// ── 10. Home ─────────────────────────────────────────────────────────────────
// Two-step home: MC_Direct sets the actual position, but does NOT raise the axis
// calibrated/Homed flag. MC_ForceCalibration then sets that flag (no motion, no
// position change). _homeCmd stays TRUE across both steps so all "home active"
// gates (jog/move blocking, fault) remain valid for the whole sequence.
IF NOT _homeCmd THEN
    _homeStep := 0;                     // sequence aborted elsewhere (stop/reset) → reset step
END_IF

// Step 1: set position
_mcHome(
    Axis       := Axis,
    Execute    := _homeCmd AND (_homeStep = 1),
    Position   := _homePosition,
    HomingMode := MC_Direct
);
IF _mcHome.Done AND (_homeStep = 1) THEN
    _homeStep          := 2;            // position set → now flag the axis as calibrated
    _dbgHomeDirectDone := TRUE;         // latch (diagnostic)
    // Retain the teach (section 10b) as an offset from the RAW encoder position, so it can be
    // re-applied after the NC restarts. Raw = the position before MC_Direct minus whatever offset
    // the running NC already applied.
    IF _retainHome THEN
        _homeOffset      := _homePosition - (_homeActAtStart - _ncOffsetApplied);
        _ncOffsetApplied := _homeOffset;
        _homeTaughtPos   := _homePosition;
        _homeTaught      := TRUE;
    END_IF
END_IF
IF _mcHome.Error THEN
    _homeCmd  := FALSE;
    _homeStep := 0;
    _lastMcErrorId := _mcHome.ErrorID;
    setFault(TRUE, CONCAT('Home error: ', UDINT_TO_STRING(_mcHome.ErrorID)));
END_IF
IF _homeStep > _dbgHomeMaxStep THEN _dbgHomeMaxStep := _homeStep; END_IF

// Step 2: set calibrated/Homed flag
_mcForceCal(
    Axis       := Axis,
    Execute    := _homeCmd AND (_homeStep = 2),
    HomingMode := MC_ForceCalibration
);
IF _mcForceCal.Done THEN
    _homeCmd        := FALSE;
    _homeStep       := 0;
    _dbgHomeCalDone := TRUE;            // latch (diagnostic)
END_IF
IF _mcForceCal.Error THEN
    _homeCmd         := FALSE;
    _homeStep        := 0;
    _dbgHomeCalError := TRUE;           // latch (diagnostic)
    _dbgHomeCalErrID := _mcForceCal.ErrorID;
    _lastMcErrorId := _mcForceCal.ErrorID;
    setFault(TRUE, CONCAT('Home cal error: ', UDINT_TO_STRING(_mcForceCal.ErrorID)));
END_IF

// ── 10b. Retained home ────────────────────────────────────────────────────────
// A taught home is kept (VAR PERSISTENT _homeTaught/_homeOffset) until the next teach — through
// PLC/NC restarts, activations and power cycles. MC_Direct only shifts the position inside the
// RUNNING NC, so after an NC restart (every activation) the axis reports the raw absolute-encoder
// position and is not homed. Once per PLC start, after the axis IO has been valid for 1 s (never
// act on a 0 read before EtherCAT is up), check the NC:
//   - not homed → the NC restarted and dropped the offset: MC_SetPosition(raw + offset), then
//                 MC_ForceCalibration. No motion and no enable needed.
//   - homed     → only the PLC restarted; the running NC still carries the offset: do nothing.
// Requires an ABSOLUTE encoder (cfgRetainHome := FALSE on an incremental one) and an NC encoder
// config that does not set the calibration flag by itself at startup.
_homeRestoreDelay(
    IN := _retainHome AND NOT _homeRestoreChecked
          AND NOT Axis.NcToPlc.StateDWord.30      // IoDataInvalid (StateDWord is a plain DWORD in Tc2_MC2)
          AND NOT Axis.NcToPlc.StateDWord.28      // DriveDeviceError
          AND NOT Axis.Status.Error,
    PT := T#1S
);
IF _homeRestoreDelay.Q THEN
    _homeRestoreChecked := TRUE;
    IF Axis.Status.Homed THEN
        _ncOffsetApplied := SEL(_homeTaught, 0.0, _homeOffset);
    ELSIF _homeTaught AND NOT _homeCmd AND NOT _externalControl THEN
        _ncOffsetApplied   := 0.0;
        _homeRestoreTarget := Axis.NcToPlc.ActPos + _homeOffset;
        _homeRestoreStep   := 1;
    END_IF
END_IF

_mcRestorePos(
    Axis     := Axis,
    Execute  := (_homeRestoreStep = 1),
    Position := _homeRestoreTarget,
    Mode     := FALSE                   // absolute
);
IF _mcRestorePos.Done AND (_homeRestoreStep = 1) THEN
    _ncOffsetApplied := _homeOffset;
    _homeRestoreStep := 2;
END_IF
IF _mcRestorePos.Error THEN
    _homeRestoreStep := 0;
    _lastMcErrorId := _mcRestorePos.ErrorID;
    setFault(TRUE, CONCAT('Home restore error: ', UDINT_TO_STRING(_mcRestorePos.ErrorID)));
END_IF

_mcRestoreCal(
    Axis       := Axis,
    Execute    := (_homeRestoreStep = 2),
    HomingMode := MC_ForceCalibration
);
IF _mcRestoreCal.Done THEN
    _homeRestoreStep := 0;
END_IF
IF _mcRestoreCal.Error THEN
    _homeRestoreStep := 0;
    _lastMcErrorId := _mcRestoreCal.ErrorID;
    setFault(TRUE, CONCAT('Home restore cal error: ', UDINT_TO_STRING(_mcRestoreCal.ErrorID)));
END_IF

// ── 11. Move execution state machine ──────────────────────────────────────────
// _moveExecState: 0=idle, 1=one-scan-abort (all Execute FALSE), 2=executing
// While yielded to an external coordinator (e.g. fb_CamCoupler), keep the state machine idle
// so every move block is driven Execute:=FALSE and never fights the external coupling.
IF _externalControl THEN
    _moveExecState := 0;
END_IF
// Arm new move request (set by cmdStart)
IF _startMoveReq AND NOT _stopCmd AND NOT _externalControl THEN
    _startMoveReq     := FALSE;
    _currentMoveIndex := _pendingIndex;
    _activeMoveMode   := _pendingMode;
    stsMoveDone       := FALSE;
    _haltCmd          := FALSE;
    _jogPositive      := FALSE;
    _jogNegative      := FALSE;
    IF _moveExecState = 2 THEN
        _moveExecState := 1; // one clear scan before rising edge on new block
    ELSE
        _moveExecState := 2;
    END_IF
END_IF

CASE _moveExecState OF

    0, 1: // Idle or abort-scan: drive all move blocks with Execute FALSE
        _mcMoveAbs(Axis := Axis, Execute := FALSE, Position := 0.0,     Velocity := 1.0, Acceleration := 1.0, Deceleration := 1.0, Jerk := 0.0);
        _mcMoveRel(Axis := Axis, Execute := FALSE, Distance := 0.0,     Velocity := 1.0, Acceleration := 1.0, Deceleration := 1.0, Jerk := 0.0);
        _mcMoveVel(Axis := Axis, Execute := FALSE);
        _mcTorque( Axis := Axis, Execute := FALSE);
        _mcMoveMod(Axis := Axis, Execute := FALSE);
        IF _moveExecState = 1 THEN
            _moveExecState := 2; // transition to executing next scan
        END_IF

    2: // Executing - drive only the active mode block; others get Execute FALSE
        CASE _activeMoveMode OF

            E_Axis_Mode.eAbsolute:
                _mcMoveAbs(
                    Axis         := Axis,
                    Execute      := TRUE,
                    Position     := moves[_currentMoveIndex].position,
                    Velocity     := moves[_currentMoveIndex].velocity,
                    Acceleration := moves[_currentMoveIndex].acceleration,
                    Deceleration := moves[_currentMoveIndex].deceleration,
                    Jerk         := moves[_currentMoveIndex].jerk
                );
                _mcMoveRel(Axis := Axis, Execute := FALSE, Distance := 0.0,     Velocity := 1.0, Acceleration := 1.0, Deceleration := 1.0, Jerk := 0.0);
                _mcMoveVel(Axis := Axis, Execute := FALSE);
                _mcTorque( Axis := Axis, Execute := FALSE);
                _mcMoveMod(Axis := Axis, Execute := FALSE);
                IF _mcMoveAbs.Done THEN
                    stsMoveDone    := TRUE;
                    _moveExecState := 0;
                END_IF
                IF _mcMoveAbs.Error THEN
                    _moveExecState := 0;
                    _lastMcErrorId := _mcMoveAbs.ErrorID;
                    setFault(TRUE, CONCAT(CONCAT('Move [', CONCAT(moves[_currentMoveIndex].moveName, '] error: ')), UDINT_TO_STRING(_mcMoveAbs.ErrorID)));
                END_IF

            E_Axis_Mode.eRelative:
                _mcMoveRel(
                    Axis         := Axis,
                    Execute      := TRUE,
                    Distance     := moves[_currentMoveIndex].position,
                    Velocity     := moves[_currentMoveIndex].velocity,
                    Acceleration := moves[_currentMoveIndex].acceleration,
                    Deceleration := moves[_currentMoveIndex].deceleration,
                    Jerk         := moves[_currentMoveIndex].jerk
                );
                _mcMoveAbs(Axis := Axis, Execute := FALSE, Position := 0.0,     Velocity := 1.0, Acceleration := 1.0, Deceleration := 1.0, Jerk := 0.0);
                _mcMoveVel(Axis := Axis, Execute := FALSE);
                _mcTorque( Axis := Axis, Execute := FALSE);
                _mcMoveMod(Axis := Axis, Execute := FALSE);
                IF _mcMoveRel.Done THEN
                    stsMoveDone    := TRUE;
                    _moveExecState := 0;
                END_IF
                IF _mcMoveRel.Error THEN
                    _moveExecState := 0;
                    _lastMcErrorId := _mcMoveRel.ErrorID;
                    setFault(TRUE, CONCAT(CONCAT('Move [', CONCAT(moves[_currentMoveIndex].moveName, '] error: ')), UDINT_TO_STRING(_mcMoveRel.ErrorID)));
                END_IF

            E_Axis_Mode.eVelocity:
                _mcMoveVel(
                    Axis         := Axis,
                    Execute      := TRUE,
                    Velocity     := moves[_currentMoveIndex].velocity,
                    Acceleration := moves[_currentMoveIndex].acceleration,
                    Deceleration := moves[_currentMoveIndex].deceleration,
                    Jerk         := moves[_currentMoveIndex].jerk,
                    Direction    := moves[_currentMoveIndex].direction
                );
                _mcMoveAbs(Axis := Axis, Execute := FALSE, Position := 0.0,     Velocity := 1.0, Acceleration := 1.0, Deceleration := 1.0, Jerk := 0.0);
                _mcMoveRel(Axis := Axis, Execute := FALSE, Distance := 0.0,     Velocity := 1.0, Acceleration := 1.0, Deceleration := 1.0, Jerk := 0.0);
                _mcTorque( Axis := Axis, Execute := FALSE);
                _mcMoveMod(Axis := Axis, Execute := FALSE);
                IF _mcMoveVel.InVelocity THEN
                    stsMoveDone := TRUE; // velocity setpoint reached; block stays active
                END_IF
                IF _mcMoveVel.Error THEN
                    _moveExecState := 0;
                    _lastMcErrorId := _mcMoveVel.ErrorID;
                    setFault(TRUE, CONCAT(CONCAT('Move [', CONCAT(moves[_currentMoveIndex].moveName, '] error: ')), UDINT_TO_STRING(_mcMoveVel.ErrorID)));
                END_IF

            E_Axis_Mode.eTorque:
                // Direction in torque mode is the SIGN of Torque (MC_TorqueControl has
                // no Direction input). moves[].direction is unused here.
                _mcTorque(
                    Axis             := Axis,
                    Execute          := TRUE,
                    ContinuousUpdate := TRUE,
                    Torque           := moves[_currentMoveIndex].torque,
                    TorqueRamp       := moves[_currentMoveIndex].torqueRamp
                );
                _mcMoveAbs(Axis := Axis, Execute := FALSE, Position := 0.0,     Velocity := 1.0, Acceleration := 1.0, Deceleration := 1.0, Jerk := 0.0);
                _mcMoveRel(Axis := Axis, Execute := FALSE, Distance := 0.0,     Velocity := 1.0, Acceleration := 1.0, Deceleration := 1.0, Jerk := 0.0);
                _mcMoveVel(Axis := Axis, Execute := FALSE);
                _mcMoveMod(Axis := Axis, Execute := FALSE);
                IF _mcTorque.InTorque THEN
                    stsMoveDone := TRUE; // torque setpoint reached; block stays active
                END_IF
                IF _mcTorque.Error THEN
                    _moveExecState := 0;
                    _lastMcErrorId := _mcTorque.ErrorID;
                    setFault(TRUE, CONCAT(CONCAT('Move [', CONCAT(moves[_currentMoveIndex].moveName, '] error: ')), UDINT_TO_STRING(_mcTorque.ErrorID)));
                END_IF
                // Software velocity limit: MC_TorqueControl has no velocity clamp and this
                // drive can't enforce one, so torque mode could run away (e.g. wire break).
                // moves[].velocity is reused as the max |velocity| permitted during torque.
                // Trip a locked MC_Stop + fault if exceeded. (Tune with margin/debounce if it
                // nuisance-trips on transients.)
                IF moves[_currentMoveIndex].velocity > 0.0
                   AND ABS(Axis.NcToPlc.ActVelo) > moves[_currentMoveIndex].velocity THEN
                    _stopCmd       := TRUE;
                    _moveExecState := 0;
                    setFault(TRUE, CONCAT('Torque velo limit: ', moves[_currentMoveIndex].moveName));
                END_IF

            E_Axis_Mode.eModulo:
                // Absolute target WITHIN one modulo period (e.g. 0..360 deg) in a FORCED direction:
                // moves[].direction = MC_Positive_Direction / MC_Negative_Direction / MC_Shortest_Way /
                // MC_Current_Direction. Unlike eAbsolute (MC_MoveAbsolute on the accumulated position,
                // which unwinds every turn back to that number), this goes to the next crossing of the
                // target in the chosen direction - "turn backwards until 0 deg". Uses the NC axis's
                // modulo factor; meant for rotary axes.
                _mcMoveMod(
                    Axis         := Axis,
                    Execute      := TRUE,
                    Position     := moves[_currentMoveIndex].position,
                    Velocity     := moves[_currentMoveIndex].velocity,
                    Acceleration := moves[_currentMoveIndex].acceleration,
                    Deceleration := moves[_currentMoveIndex].deceleration,
                    Jerk         := moves[_currentMoveIndex].jerk,
                    Direction    := moves[_currentMoveIndex].direction
                );
                _mcMoveAbs(Axis := Axis, Execute := FALSE, Position := 0.0,     Velocity := 1.0, Acceleration := 1.0, Deceleration := 1.0, Jerk := 0.0);
                _mcMoveRel(Axis := Axis, Execute := FALSE, Distance := 0.0,     Velocity := 1.0, Acceleration := 1.0, Deceleration := 1.0, Jerk := 0.0);
                _mcMoveVel(Axis := Axis, Execute := FALSE);
                _mcTorque( Axis := Axis, Execute := FALSE);
                IF _mcMoveMod.Done THEN
                    stsMoveDone    := TRUE;
                    _moveExecState := 0;
                END_IF
                IF _mcMoveMod.Error THEN
                    _moveExecState := 0;
                    _lastMcErrorId := _mcMoveMod.ErrorID;
                    setFault(TRUE, CONCAT(CONCAT('Move [', CONCAT(moves[_currentMoveIndex].moveName, '] error: ')), UDINT_TO_STRING(_mcMoveMod.ErrorID)));
                END_IF

        ELSE
            // A mode with no implementation (eHalt/eStop/eHome/eSetPosition/eExternal as a move)
            // used to sit in _moveExecState = 2 forever with no MC block running and stsMoveDone
            // never TRUE - a sequence waiting on it would hang. Refuse it loudly instead.
            _moveExecState := 0;
            setFault(TRUE, CONCAT(CONCAT('Move [', CONCAT(moves[_currentMoveIndex].moveName, '] mode not supported: ')), INT_TO_STRING(_activeMoveMode)));

        END_CASE

        // Overtorque limit: fault if |actual torque| exceeds this move's configured limit
        // during execution. Unlike the torque-mode velocity watchdog (above), this applies to
        // EVERY mode — a jam/collision on a position or velocity move shows up as excess torque
        // just as on a torque move. moves[].cfgTorqueLimit = 0 disables the check. Trip → locked
        // MC_Stop + fault (cmdReset required), matching the velocity watchdog. Guarded on
        // _moveExecState = 2 so a move that just completed/errored this scan can't also trip.
        // (Add a debounce TON here if it nuisance-trips on accel transients.)
        IF _moveExecState = 2
           AND moves[_currentMoveIndex].cfgTorqueLimit > 0.0
           AND ABS(Axis.NcToPlc.ActTorque) > moves[_currentMoveIndex].cfgTorqueLimit THEN
            _stopCmd       := TRUE;
            _moveExecState := 0;
            setFault(TRUE, CONCAT('Overtorque limit: ', moves[_currentMoveIndex].moveName));
        END_IF

END_CASE

// ── 12. Jog ──────────────────────────────────────────────────────────────────
// Level-triggered: hold = continuous jog. Requires axis interlock met (req. 4).
// Effective jog dynamics: when the pendant owns the jog it supplies its own speed/accel
// (falling back to the configured jog values if <= 0); HMI jog always uses the configured
// values. Computed here so the pendant never overwrites the HMI's configured _jogVelocity.
_jogVeloEff  := _jogVelocity;
_jogAccelEff := _jogAccel;
IF _jogSource = E_Axis_JogSource.ePendant THEN
    IF inpPendantJogVelo  > 0.0 THEN _jogVeloEff  := inpPendantJogVelo;  END_IF
    IF inpPendantJogAccel > 0.0 THEN _jogAccelEff := inpPendantJogAccel; END_IF
END_IF
// Clamp to the NC axis's maximum velocity. A jog above it is refused by the NC (MC_Jog error
// 0x4221 'velocity not allowed') and the axis simply does not move - an operator jog speed of
// 80 mm/s on a 27.3 mm/s axis made HMI jog look dead. stsJogVelocity shows the clamped value.
// (MC_ReadParameter AxisVeloMax answers ADS 0x701 'service not supported' - read the whole set.)
_readParamsRetry(IN := (_ncMaxVelocity <= 0.0) AND NOT _readParamsExec, PT := T#2S);
IF _readParamsRetry.Q THEN
    _readParamsExec := TRUE;
END_IF
_mcReadParams(Parameter := _axisParams, Axis := Axis, Execute := _readParamsExec);
IF _mcReadParams.Done THEN
    _readParamsExec := FALSE;
    IF _axisParams.fVeloMaximum > 0.0 THEN
        _ncMaxVelocity := _axisParams.fVeloMaximum;
    END_IF
ELSIF _mcReadParams.Error THEN
    _readParamsExec := FALSE;   // retried by _readParamsRetry
END_IF
IF _ncMaxVelocity > 0.0 AND _jogVeloEff > _ncMaxVelocity THEN
    _jogVeloEff := _ncMaxVelocity;
END_IF
// Pendant deflection as a FRACTION of the clamped speed: scaling before the clamp saturated
// (configured 80 mm/s on a 27.3 mm/s axis -> anything past a third of the stick was full speed).
IF _jogSource = E_Axis_JogSource.ePendant AND inpPendantJogFraction > 0.0 THEN
    _jogVeloEff := _jogVeloEff * LIMIT(0.0, inpPendantJogFraction, 1.0);
END_IF

_pjGate := _mcPower.Status AND Interlock.outInterlockOK AND NOT stsFaulted AND NOT _stopCmd AND NOT _homeCmd
           AND NOT _torqueJogEngaged AND (_moveExecState = 0) AND NOT _externalControl AND NOT _jogGotoBusy;

_mcJog(
    Axis         := Axis,
    Mode         := MC_JOGMODE_CONTINOUS,
    JogForward   := _jogPositive AND _jogSource <> E_Axis_JogSource.ePendant AND NOT _externalControl AND NOT _jogGotoBusy AND _mcPower.Status AND Interlock.outInterlockOK AND NOT stsFaulted AND NOT _stopCmd AND NOT _homeCmd AND NOT _torqueJogEngaged AND (_moveExecState = 0),
    JogBackwards := _jogNegative AND _jogSource <> E_Axis_JogSource.ePendant AND NOT _externalControl AND NOT _jogGotoBusy AND _mcPower.Status AND Interlock.outInterlockOK AND NOT stsFaulted AND NOT _stopCmd AND NOT _homeCmd AND NOT _torqueJogEngaged AND (_moveExecState = 0),
    Velocity     := _jogVeloEff,
    Acceleration := _jogAccelEff
);
// A refused jog used to be silent (the axis just did not move) - report it.
_jogErrorEdge(CLK := _mcJog.Error);
IF _jogErrorEdge.Q THEN
    _lastMcErrorId := _mcJog.ErrorID;
    setFault(TRUE, CONCAT('Jog error: ', UDINT_TO_STRING(_mcJog.ErrorID)));
END_IF

// ── 12b. Pendant jog ──────────────────────────────────────────────────────────
// MC_MoveVelocity at _jogVeloEff, which follows the stick / speed modifier live. Tc2_MC2
// MC_MoveVelocity takes a new speed only on a rising Execute, so a change of more than 2 % (at
// most every 20 ms) drops Execute for one scan and re-triggers it - the NC blends to the new
// speed. A direction change re-triggers too (the NC reverses through zero). Release (stick in
// its dead zone, dead-man let go, pendant deselected) or the gate dropping -> MC_Halt at the jog
// accel, held until standstill. MC_Stop (stop / fault / STO) supersedes it: no halt is issued
// while _stopCmd, and power-off needs none.
_pjDir := 0;
IF _jogSource = E_Axis_JogSource.ePendant AND _pjGate AND _jogVeloEff > 0.0 THEN
    IF _jogPositive THEN
        _pjDir := 1;
    ELSIF _jogNegative THEN
        _pjDir := -1;
    END_IF
END_IF
IF _pjDir <> 0 AND _pjDir = _pjDirPrev THEN
    IF _pjVelExec AND _pjRetrig.Q AND ABS(_jogVeloEff - _pjVeloSent) > 0.02 * MAX(_jogVeloEff, _pjVeloSent) THEN
        _pjVelExec := FALSE;
    ELSIF NOT _pjVelExec THEN
        _pjVelExec  := TRUE;
        _pjVeloSent := _jogVeloEff;
        _pjMoving   := TRUE;
    END_IF
ELSE
    _pjVelExec := FALSE;
END_IF
_pjDirPrev := _pjDir;
IF _stopCmd OR NOT _mcPower.Status THEN
    _pjMoving := FALSE;     // MC_Stop / power-off own the axis now
END_IF
_pjRetrig(IN := _pjVelExec, PT := T#20MS);
_mcPendantVel(
    Axis         := Axis,
    Execute      := _pjVelExec,
    Velocity     := _pjVeloSent,
    Acceleration := _jogAccelEff,
    Deceleration := _jogAccelEff,
    Jerk         := 0.0,
    Direction    := SEL(_pjDir > 0, MC_Negative_Direction, MC_Positive_Direction)
);
_mcPendantHalt(
    Axis         := Axis,
    Execute      := _pjMoving AND _pjDir = 0,
    Deceleration := _jogAccelEff,
    Jerk         := 0.0
);
IF _mcPendantHalt.Done OR _mcPendantHalt.Error OR _mcPendantHalt.CommandAborted THEN
    _pjMoving := FALSE;
END_IF
_pjErrorEdge(CLK := _mcPendantVel.Error);
IF _pjErrorEdge.Q THEN
    _lastMcErrorId := _mcPendantVel.ErrorID;
    setFault(TRUE, CONCAT('Pendant jog error: ', UDINT_TO_STRING(_mcPendantVel.ErrorID)));
END_IF

// Overtorque limit for position jog: global analogue of the per-move cfgTorqueLimit.
// While jogging, trip a locked MC_Stop + fault if |actual torque| exceeds _jogTorqueLimit
// (0 = disabled). Excludes torque-jog, which deliberately commands torque and is bounded by
// its own _torqueJogMaxLimit clamp. MC_Stop reacts next scan (same 1-scan latency as the
// STO / interlock-loss trips), and clearing the jog flags stops MC_Jog commanding.
IF (_jogPositive OR _jogNegative)
   AND _jogTorqueLimit > 0.0
   AND ABS(Axis.NcToPlc.ActTorque) > _jogTorqueLimit THEN
    _jogPositive := FALSE;
    _jogNegative := FALSE;
    _stopCmd     := TRUE;
    IF NOT stsFaulted THEN
        setFault(TRUE, 'Overtorque limit: jog');
    END_IF
END_IF

// ── 12b. Torque jog (dead-man interactive torque) ─────────────────────────────
// Engage on first press (while powered/safe/idle). Stay engaged while held OR until the
// released torque has ramped back to ~0, so letting go RAMPS down instead of snapping.
// Held → command the entered torque; released → command 0.0 (ramps at _torqueJogRamp).
// Ends FREE at 0 torque, axis stays enabled — no MC_Stop, so no NC 0x4268. A max-velocity
// trip cuts the torque command (ramps to 0) if the axis runs away, since torque control has
// no speed clamp of its own. NOT safety-rated — the PLC interlocks/STO are.
IF _torqueJogActive AND NOT _jogGotoBusy AND _mcPower.Status AND Interlock.outInterlockOK AND NOT stsFaulted AND NOT _stopCmd THEN
    _torqueJogEngaged := TRUE;
END_IF
// Torque-jog overspeed trip [unit/s], 0 = disabled. PERSISTENT: the operator's value is
// retained across PLC restart (backed by VAR PERSISTENT _tjMaxVel). On the first scan after
// a (re)start, push the retained value OUT to the HMI field so the HMI shows it instead of
// clobbering it with its power-up 0; from then on the HMI field is the live editor and its
// value (including 0 = disable) is copied back into the persistent store. Assumes the HMI
// reads the seeded value on (re)connect rather than immediately re-writing a cached one.
IF NOT _tjMaxVelInit THEN
    HMI.Commands.ocmdTorqueJogMaxVel := _tjMaxVel;   // seed HMI from retained value
    _tjMaxVelInit := TRUE;
ELSE
    _tjMaxVel := HMI.Commands.ocmdTorqueJogMaxVel;   // operator edits → persist
END_IF
IF _torqueJogEngaged AND _tjMaxVel > 0.0 AND ABS(Axis.NcToPlc.ActVelo) > _tjMaxVel THEN
    _torqueJogActive := FALSE;   // overspeed → stop commanding torque (ramp to 0)
    setFault(TRUE, 'Torque-jog overspeed');
END_IF
_mcTorqueJog(
    Axis             := Axis,
    Execute          := _torqueJogEngaged AND NOT _externalControl AND NOT _jogGotoBusy AND _mcPower.Status AND Interlock.outInterlockOK AND NOT stsFaulted AND NOT _stopCmd,
    ContinuousUpdate := TRUE,
    Torque           := SEL(_torqueJogActive, 0.0, _torqueJogValue),   // held → value; released → 0
    TorqueRamp       := _torqueJogRamp
);
// Release complete: not held and torque back to ~0 → disengage (drop Execute; drive holds 0/free).
IF _torqueJogEngaged AND NOT _torqueJogActive AND ABS(Axis.NcToPlc.ActTorque) < _stopTorqueThreshold THEN
    _torqueJogEngaged := FALSE;
END_IF

// ── 12c. Position jog ("go to position") ──────────────────────────────────────
// Discrete absolute move to an operator-entered target (angle or mm) at the jog velocity/accel -
// a jog subvariant selected on the HMI. Started by cmdJogGoto (via ocmdJogGoto). Mutually exclusive
// with speed-jog / torque-jog / configured moves / home (gated here and in cmdJogGoto). Same safety
// chain as jog: a stop / fault / STO / interlock loss aborts it via MC_Stop and clears _jogGotoBusy.
// For a modulo axis this goes to the absolute target; shortest-path would use MC_MoveModulo (future).
_mcJogGoto(
    Axis         := Axis,
    Execute      := _jogGotoBusy AND NOT _externalControl AND _mcPower.Status AND Interlock.outInterlockOK
                    AND NOT stsFaulted AND NOT _stopCmd AND NOT _homeCmd AND (_moveExecState = 0)
                    AND NOT _jogPositive AND NOT _jogNegative AND NOT _torqueJogEngaged,
    Position     := _jogGotoTarget,
    Velocity     := _jogVeloEff,
    Acceleration := _jogAccelEff,
    Deceleration := _jogAccelEff,
    Jerk         := 0.0
);
IF _mcJogGoto.Done THEN
    _jogGotoBusy := FALSE;               // reached target
END_IF
IF _mcJogGoto.CommandAborted THEN
    _jogGotoBusy := FALSE;               // superseded by a stop / other command
END_IF
IF _mcJogGoto.Error THEN
    _jogGotoBusy := FALSE;
    _lastMcErrorId := _mcJogGoto.ErrorID;
    setFault(TRUE, CONCAT('Jog goto error: ', UDINT_TO_STRING(_mcJogGoto.ErrorID)));
END_IF

// ── 13. Velocity override (local or global) ──────────────────────────────────
// Effective velocity override = the machine-global value when inpGlobalOverrideEnable is set,
// otherwise the axis-local _velocityOverride (set from HMI). The global INT [%] is clamped to
// 0..100 (0 = axis held at 0%). Only the effective value is applied and reported. AccFactor
// always tracks the local accel override.
// VelFactor and AccFactor are 0.0 to 1.0 (MC_SetOverride convention).
IF inpGlobalOverrideEnable THEN
    _activeVelocityOverride := LIMIT(0.0, INT_TO_LREAL(inpGlobalOverride), 100.0);
ELSE
    _activeVelocityOverride := _velocityOverride;
END_IF
_mcOverride(
    Axis      := Axis,
    Enable    := _isEnabled,
    VelFactor := _activeVelocityOverride / 100.0,
    AccFactor := _accelOverride / 100.0
);

// ── 14. NC-level axis error detection ────────────────────────────────────────
IF Axis.Status.Error AND NOT stsFaulted THEN
    setFault(TRUE, CONCAT('Axis error: ', UDINT_TO_STRING(Axis.NcToPlc.ErrorCode)));
END_IF

// ── 15. Status outputs ───────────────────────────────────────────────────────
stsEnabled    := _mcPower.Status;
stsMoving     := Axis.Status.DiscreteMotion OR Axis.Status.ContinuousMotion;
stsStandstill := Axis.Status.Standstill;
stsInTarget   := Axis.Status.InTargetPosition;
stsCurrentMove:= _currentMoveIndex;

// ── 16. HMI status update ────────────────────────────────────────────────────
// Inherited base-device HMI values (deviceName, enabled, stsInAuto, fault, interlock).
// DeviceLogic() filled the inherited HMIbaseDevice VAR at the top of this scan.
HMI.HMIbaseDevice              := HMIbaseDevice;
HMI.Status.stsEnabled          := stsEnabled;
HMI.Status.stsHomed            := Axis.Status.Homed;       // referenced/calibrated
HMI.Status.stsStandstill       := stsStandstill;
HMI.Status.stsMoving           := stsMoving;
HMI.Status.stsInTargetPos      := stsInTarget;
HMI.Status.stsError            := Axis.Status.Error;
// The NC axis error, else the last motion-block error (a refused jog/move is an MC_* FB error, not an
// axis error) - so the HMI's TwinCAT NC lookup can describe it. Cleared by cmdReset.
HMI.Status.stsErrorID          := SEL(Axis.NcToPlc.ErrorCode <> 0, _lastMcErrorId, Axis.NcToPlc.ErrorCode);
// Full AXIS_REF.Status snapshot - exposes every status flag this lib version has
HMI.Status.stsAxisStatus       := Axis.Status;
// Live process values → outputs (single source), then mirror into HMI.Status.
stsActualPosition := Axis.NcToPlc.ActPos;
stsActualVelocity := Axis.NcToPlc.ActVelo;
stsNcMaxVelocity  := _ncMaxVelocity;     // what the jog clamp uses - also lets callers size their own commands
stsActualTorque   := Axis.NcToPlc.ActTorque;   // actual torque from drive
HMI.Status.stsActualPosition   := stsActualPosition;
HMI.Status.stsActualVelocity   := stsActualVelocity;
HMI.Status.stsActualTorque     := stsActualTorque;
// Modulo position: NC-computed, wrapped into one period. Always populated; the HMI shows it
// instead of stsActualPosition only when stsIsModulo (set below). ActPos above is un-wrapped.
HMI.Status.stsModuloActPos     := Axis.NcToPlc.ModuloActPos;
HMI.Status.stsModuloActTurns   := Axis.NcToPlc.ModuloActTurns;
// Setpoints → outputs (single source), then mirror into HMI.Status.
stsSetPosition := Axis.NcToPlc.SetPos;
stsSetVelocity := Axis.NcToPlc.SetVelo;
// Commanded torque — no NC setpoint exists; report what the FB is feeding the drive.
IF _torqueJogEngaged THEN
    stsSetTorque := SEL(_torqueJogActive, 0.0, _torqueJogValue);          // held → value, releasing → 0
ELSIF _moveExecState = 2 AND _activeMoveMode = E_Axis_Mode.eTorque THEN
    stsSetTorque := moves[_currentMoveIndex].torque;                       // active torque move
ELSE
    stsSetTorque := 0.0;                                                   // idle / non-torque
END_IF
HMI.Status.stsSetPosition      := stsSetPosition;
HMI.Status.stsSetVelocity      := stsSetVelocity;
HMI.Status.stsSetTorque        := stsSetTorque;
HMI.Status.stsFollowingError   := Axis.NcToPlc.SetPos - Axis.NcToPlc.ActPos;
HMI.Status.stsHomeBusy         := _homeCmd;                              // whole 2-step sequence in progress
HMI.Status.stsHomeDone         := _mcForceCal.Done;                      // sequence complete = calibrated flag set
HMI.Status.stsHomeError        := _mcHome.Error OR _mcForceCal.Error;
HMI.Status.stsHomeErrorID      := SEL(_mcForceCal.Error, _mcHome.ErrorID, _mcForceCal.ErrorID);
HMI.Status.stsHomePosition     := _homePosition;
HMI.Status.stsCurrentMoveIndex := _currentMoveIndex;
IF _currentMoveIndex >= 1 AND _currentMoveIndex <= 20 THEN
    HMI.Status.stsCurrentMoveName := moves[_currentMoveIndex].moveName;
ELSE
    HMI.Status.stsCurrentMoveName := '';
END_IF
HMI.Status.stsSelectedMove     := _selectedMove;
HMI.Status.stsConfirmPending   := _confirmPending;
HMI.Status.stsMoveConfigLoaded     := _hmiMoveConfigLoaded;
HMI.Status.stsMoveConfigApplyError := _moveConfigApplyError;
HMI.Status.stsMoveConfigErrorText  := _moveConfigErrorText;
HMI.Status.stsMoveDone         := stsMoveDone;
HMI.Status.stsMoveBusy         := (_moveExecState = 2);
HMI.Status.stsActiveMoveMode   := _activeMoveMode;
HMI.Status.stsExternalControl  := _externalControl;
HMI.Status.stsAxisType         := _axisType;
HMI.Status.stsUnit             := _unit;
HMI.Status.stsIsModulo         := _isModulo;
HMI.Status.stsVelocityOverride     := _activeVelocityOverride;   // effective: global if active, else local
HMI.Status.stsGlobalOverrideActive := inpGlobalOverrideEnable;
HMI.Status.stsJogVelocity      := _jogVeloEff;   // effective (pendant speed when it owns, else configured)
HMI.Status.stsJogAcceleration  := _jogAccelEff;
HMI.Status.stsJogSource        := _jogSource;    // none / HMI / pendant (which input owns the jog)
HMI.Status.stsPendantMode      := inpPendantMode OR inpPendantEnable;   // pendant owns the jog - HMI jog locked out
HMI.Status.stsPendantDeadman   := inpPendantEnable;                     // dead-man held - pendant can move the axis
HMI.Status.stsHomeRetained     := _homeTaught AND _retainHome;          // a taught home is stored and survives restarts
HMI.Status.stsJogTorqueLimit   := _jogTorqueLimit;
HMI.Status.stsTorqueJogActive  := _torqueJogEngaged;
HMI.Status.stsTorqueJogMaxVel  := _tjMaxVel;
HMI.Status.stsJogGotoBusy      := _jogGotoBusy;
HMI.Status.stsJogGotoDone      := _mcJogGoto.Done;
HMI.Status.stsJogGotoPos       := _jogGotoTarget;
HMI.Status.stsSTO              := inpSTO;
HMI.Status.stsSafetyInhibited  := NOT inpSTO;   // motion inhibited by safety (STO active) - not a fault
FOR _i := 1 TO 20 DO
    HMI.Status.moves[_i]          := moves[_i];
    HMI.Status.moveInterlocks[_i] := _moveInterlocks[_i].getHMIdata();
END_FOR

// Execute a pre-defined move by index (1-20).
// Checks axis-level interlock then move-level interlock before arming.
// Fault description format: "I_NOK: <description>" or "Move I_NOK: <description>"
METHOD PUBLIC cmdStart : BOOL
VAR_INPUT
    moveIndex : INT;  // 1-20
END_VAR
IF moveIndex < 1 OR moveIndex > 20 THEN
    RETURN;
END_IF

// Yielded to a coordinator - reject quietly. Do NOT setFault: a fault gates MC_Power (section 6)
// and would drop the axis and break any active cam coupling.
IF _externalControl THEN
    cmdStart := FALSE;
    RETURN;
END_IF

IF NOT _mcPower.Status THEN
    setFault(TRUE, 'Axis not enabled');
    RETURN;
END_IF

IF _homeCmd THEN
    setFault(TRUE, 'Home active');
    RETURN;
END_IF

IF _jogPositive OR _jogNegative THEN
    setFault(TRUE, 'Cannot start move while jogging');
    RETURN;
END_IF

IF _torqueJogEngaged THEN
    setFault(TRUE, 'Cannot start move while torque-jogging');
    RETURN;
END_IF

IF _jogGotoBusy THEN
    setFault(TRUE, 'Cannot start move while going to position');
    RETURN;
END_IF

IF NOT Interlock.outInterlockOK THEN
    setFault(TRUE, CONCAT('I_NOK: ', Interlock.stsFirstOut));
    RETURN;
END_IF

// Re-evaluate this move's interlock immediately (also runs in main body each scan)
_moveInterlocks[moveIndex](inpConfig := moves[moveIndex].interlock);
IF NOT _moveInterlocks[moveIndex].outInterlockOK THEN
    setFault(TRUE, CONCAT('Move I_NOK: ', _moveInterlocks[moveIndex].stsFirstOut));
    RETURN;
END_IF

_pendingIndex := moveIndex;
_pendingMode  := moves[moveIndex].mode;
_startMoveReq := TRUE;
cmdStart      := TRUE;
END_METHOD

// Assign the axis home/reference position using MC_Home with HomingMode := MC_Direct.
// This does not move the axis. It is accepted only while powered, safe, and idle.
METHOD PUBLIC cmdHome : BOOL
VAR_INPUT
    homePosition : LREAL; // [unit]
END_VAR
// Yielded to a coordinator - reject quietly (a fault would drop power and break any coupling).
IF _externalControl THEN
    cmdHome := FALSE;
    RETURN;
END_IF

IF NOT _mcPower.Status THEN
    setFault(TRUE, 'Axis not enabled');
    RETURN;
END_IF

IF _stopCmd THEN
    setFault(TRUE, 'Stop active - reset required before homing');
    RETURN;
END_IF

IF stsFaulted THEN
    RETURN;
END_IF

IF NOT Interlock.outInterlockOK THEN
    setFault(TRUE, CONCAT('I_NOK: ', Interlock.stsFirstOut));
    RETURN;
END_IF

IF _moveExecState <> 0 OR _jogGotoBusy OR Axis.Status.DiscreteMotion OR Axis.Status.ContinuousMotion OR Axis.Status.Stopping THEN
    setFault(TRUE, 'Cannot home while axis is active');
    RETURN;
END_IF

// The retained home is being re-applied (a few scans after start) - reject quietly; teach again after.
IF _homeRestoreStep <> 0 THEN
    RETURN;
END_IF

// Teaching before the once-per-start retained-home check ran: settle what offset the running NC
// carries now (same rule as section 10b) so the new offset is computed from the true raw position.
// Reads the FB's own per-scan copies (HMI.Status.stsHomed, stsActualPosition), not Axis: no new
// VAR_IN_OUT access from a method (C0371), and teaching is at standstill, so last scan's value is exact.
IF NOT _homeRestoreChecked THEN
    _homeRestoreChecked := TRUE;
    _ncOffsetApplied    := SEL(HMI.Status.stsHomed AND _homeTaught, 0.0, _homeOffset);
END_IF
_homeActAtStart := stsActualPosition;

_jogPositive      := FALSE;
_jogNegative      := FALSE;
_startMoveReq     := FALSE;
_selectedMove     := 0;
_confirmPending   := FALSE;
_currentMoveIndex := 0;
_homePosition     := homePosition;
_homeCmd          := TRUE;
_homeStep         := 1;             // start at step 1 (MC_Direct set position)
// reset home diagnostics for this run
_dbgHomeMaxStep    := 0;
_dbgHomeDirectDone := FALSE;
_dbgHomeCalDone    := FALSE;
_dbgHomeCalError   := FALSE;
_dbgHomeCalErrID   := 0;
stsMoveDone       := FALSE;
cmdHome           := TRUE;
END_METHOD

// Power on the axis. Blocked if axis-level interlock not met.
METHOD PUBLIC cmdEnable : BOOL
IF NOT inpSTO THEN
    // STO active is a soft safety inhibit (see section 4), not a fault. Reject the enable
    // quietly; stsSafetyInhibited tells the operator why. Enable succeeds once STO is restored.
    cmdEnable := FALSE;
    RETURN;
END_IF

IF NOT Interlock.outInterlockOK THEN
    setFault(TRUE, CONCAT('I_NOK: ', Interlock.stsFirstOut));
    cmdEnable := FALSE;
    RETURN;
END_IF

_isEnabled := TRUE;
cmdEnable  := TRUE;
END_METHOD

// Power off the axis. Clears jog and pending moves.
METHOD PUBLIC cmdDisable : BOOL
_isEnabled     := FALSE;
_jogPositive   := FALSE;
_jogNegative   := FALSE;
_homeCmd       := FALSE;
_startMoveReq  := FALSE;
_jogGotoBusy   := FALSE;
_moveExecState := 0;
cmdDisable     := TRUE;
END_METHOD

// Forced standstill via MC_Stop. Axis stays locked until cmdReset is called.
// Immediate for every case (idle, jog, position/velocity/torque move, already stopping).
// NOTE: for a torque (CST) move this locks the axis into position hold while it was
// applying torque; to instead release a torque hold cleanly, DISABLE the axis
// (cmdDisable → MC_Power off drops torque). A graceful zero-then-stop was prototyped and
// abandoned (couldn't reliably exit CST mode — NC 0x4268, setpoint generator inactive).
METHOD PUBLIC cmdStop : BOOL
_jogPositive   := FALSE;
_jogNegative   := FALSE;
_homeCmd       := FALSE;
_startMoveReq  := FALSE;
_jogGotoBusy   := FALSE;

_stopCmd       := TRUE;
_haltCmd       := FALSE;
_moveExecState := 0;
cmdStop        := TRUE;
END_METHOD

// Interruptible stop via MC_Halt. Clears automatically when standstill reached.
// A new cmdStart can resume motion after halt completes.
METHOD PUBLIC cmdHalt : BOOL
_haltCmd       := TRUE;
_jogPositive   := FALSE;
_jogNegative   := FALSE;
_homeCmd       := FALSE;
_startMoveReq  := FALSE;
_jogGotoBusy   := FALSE;
_moveExecState := 0;
cmdHalt        := TRUE;
END_METHOD

// Clear PLC fault, release MC_Stop, trigger MC_Reset for NC errors.
// Called automatically by DeviceLogic when inpReset (machine reset) is TRUE.
METHOD cmdReset : BOOL
setFault(FALSE, '');
_stopCmd          := FALSE;
_haltCmd          := FALSE;
_resetCmd         := TRUE;
_homeCmd          := FALSE;
_startMoveReq     := FALSE;
_jogGotoBusy      := FALSE;
_moveExecState    := 0;
stsMoveDone       := FALSE;
_selectedMove     := 0;
_confirmPending   := FALSE;
_currentMoveIndex := 0;
_lastMcErrorId    := 0;
cmdReset          := TRUE;
END_METHOD

// Start positive-direction jog. Requires axis interlock met (enforced in main body).
// Level: call once, axis jogs until cmdJogStop or button released from HMI.
METHOD PUBLIC cmdJogPositive : BOOL
VAR_INPUT
    velocity    : LREAL;    // [unit/s]  - 0 = use cfgJogVelocity
    acceleration: LREAL;    // [unit/s²] - 0 = use cfgJogAcceleration
END_VAR
IF _homeCmd OR _moveExecState <> 0 OR _externalControl OR _jogGotoBusy THEN
    RETURN;
END_IF

IF velocity     > 0.0 THEN _jogVelocity := velocity;     END_IF
IF acceleration > 0.0 THEN _jogAccel    := acceleration; END_IF
_jogPositive    := TRUE;
_jogNegative    := FALSE;
cmdJogPositive  := TRUE;
END_METHOD

// Start negative-direction jog. Requires axis interlock met (enforced in main body).
METHOD PUBLIC cmdJogNegative : BOOL
VAR_INPUT
    velocity    : LREAL;    // [unit/s]  - 0 = use cfgJogVelocity
    acceleration: LREAL;    // [unit/s²] - 0 = use cfgJogAcceleration
END_VAR
IF _homeCmd OR _moveExecState <> 0 OR _externalControl OR _jogGotoBusy THEN
    RETURN;
END_IF

IF velocity     > 0.0 THEN _jogVelocity := velocity;     END_IF
IF acceleration > 0.0 THEN _jogAccel    := acceleration; END_IF
_jogNegative    := TRUE;
_jogPositive    := FALSE;
cmdJogNegative  := TRUE;
END_METHOD

// Stop jog. Axis decelerates via MC_Jog's internal decel (drive default).
METHOD PUBLIC cmdJogStop : BOOL
_jogPositive := FALSE;
_jogNegative := FALSE;
cmdJogStop   := TRUE;
END_METHOD

// Position jog: "go to position". A discrete absolute move to an operator-entered target
// (angle or mm) at the jog velocity/accel - the third jog subvariant (speed / torque / position).
// Started from the HMI via ocmdJogGoto + ocmdJogGotoPos; executed by _mcJogGoto in section 12c.
// Rejects QUIETLY (no fault) if not idle/safe, consistent with the other cmdJog* methods.
METHOD PUBLIC cmdJogGoto : BOOL
VAR_INPUT
    position : LREAL;   // [unit] absolute target (angle or mm)
END_VAR
IF _homeCmd OR _moveExecState <> 0 OR _externalControl
   OR _jogPositive OR _jogNegative OR _torqueJogEngaged OR _jogGotoBusy
   OR _stopCmd OR stsFaulted OR NOT _mcPower.Status OR NOT Interlock.outInterlockOK THEN
    RETURN;
END_IF

_jogGotoTarget := position;
_jogGotoBusy   := TRUE;
cmdJogGoto     := TRUE;
END_METHOD

// Yield axis to an external coordinator (camming/gearing layer, e.g. fb_CamCoupler).
// On enable, an interruptible cmdHalt() brings the axis to rest before the coordinator takes over.
// While yielded (_externalControl): MC_Power / MC_Reset / MC_SetOverride / status keep running so the
// axis stays powered and reportable, but ALL of the FB's own motion is suppressed - moves, jog,
// pendant jog, torque-jog and home are gated off in the scan body, and cmdStart/cmdHome/cmdJog*
// reject QUIETLY (never setFault: a fault gates MC_Power and would drop the coupling). This lets the
// coordinator command the shared AXIS_REF (MC_CamIn, etc.) without fighting the FB.
// Clearing external control does NOT re-enable motion - call cmdStart or cmdJog explicitly.
METHOD PUBLIC cmdSetExternalControl : BOOL
VAR_INPUT
    enable : BOOL;
END_VAR
_externalControl := enable;
IF enable THEN
    cmdHalt(); // interruptible stop before yielding
END_IF
cmdSetExternalControl := TRUE;
END_METHOD

// Return the full HMI interface struct for linking to an HMI symbol.
METHOD PUBLIC getHMIdata : ST_Axis_HMI_Interface
getHMIdata := HMI;
END_METHOD

METHOD FB_Init : BOOL
VAR_INPUT
    bInitRetains        : BOOL;
    bInCopyCode         : BOOL;
    cfgDeviceName       : STRING;
    cfgEnable           : BOOL;
    cfgInitEventClass   : BOOL;
    cfgJogVelocity      : LREAL;    // [unit/s]
    cfgJogAcceleration  : LREAL;    // [unit/s²]
    cfgStopDecel        : LREAL;    // [unit/s²] decel for MC_Stop
    cfgHaltDecel        : LREAL;    // [unit/s²] decel for MC_Halt
    cfgAxisType         : E_Axis_UnitType;  // eLinear / eRotary (HMI unit display)
    cfgUnit             : STRING;   // position unit label ('mm','deg',...); '' = keep default 'mm'
    cfgIsModulo         : BOOL;     // TRUE = NC axis is modulo; HMI shows modulo position (ModuloActPos)
END_VAR
THIS^.cfgDeviceName     := cfgDeviceName;
THIS^.cfgEnable         := cfgEnable;
THIS^.cfgInitEventClass := cfgInitEventClass;
IF cfgJogVelocity     > 0.0 THEN _jogVelocity := cfgJogVelocity;     END_IF
IF cfgJogAcceleration > 0.0 THEN _jogAccel    := cfgJogAcceleration; END_IF
IF cfgStopDecel       > 0.0 THEN _stopDecel   := cfgStopDecel;       END_IF
IF cfgHaltDecel       > 0.0 THEN _haltDecel   := cfgHaltDecel;       END_IF
_axisType := cfgAxisType;
IF cfgUnit <> '' THEN _unit := cfgUnit; END_IF
_isModulo := cfgIsModulo;
END_METHOD

PROPERTY PUBLIC cfgJogVelocity : LREAL
GET
cfgJogVelocity := _jogVelocity;
END_GET
SET
IF cfgJogVelocity > 0.0 THEN _jogVelocity := cfgJogVelocity; END_IF
END_SET
END_PROPERTY

PROPERTY PUBLIC cfgJogAcceleration : LREAL
GET
cfgJogAcceleration := _jogAccel;
END_GET
SET
IF cfgJogAcceleration > 0.0 THEN _jogAccel := cfgJogAcceleration; END_IF
END_SET
END_PROPERTY

// TRUE (default) = a taught home is kept until the next teach and re-applied after every NC
// restart (section 10b). Requires an ABSOLUTE encoder - set FALSE for an incremental one, whose
// raw position after a restart is meaningless. FALSE also stops recording new teaches.
PROPERTY PUBLIC cfgRetainHome : BOOL
GET
cfgRetainHome := _retainHome;
END_GET
SET
_retainHome := cfgRetainHome;
END_SET
END_PROPERTY

// [Nm or %] global overtorque trip during position jog. If |actual torque| exceeds
// this while jogging, the axis faults ('Overtorque limit: jog') and locks via MC_Stop
// (cmdReset required). 0 disables the check. Same units as Axis.NcToPlc.ActTorque.
// Does not affect torque-jog, which is bounded by its own clamp.
PROPERTY PUBLIC cfgJogTorqueLimit : LREAL
GET
cfgJogTorqueLimit := _jogTorqueLimit;
END_GET
SET
// >= 0: a value of 0 is valid and disables the trip.
IF cfgJogTorqueLimit >= 0.0 THEN _jogTorqueLimit := cfgJogTorqueLimit; END_IF
END_SET
END_PROPERTY

PROPERTY PUBLIC cfgStopDecel : LREAL
GET
cfgStopDecel := _stopDecel;
END_GET
SET
IF cfgStopDecel > 0.0 THEN _stopDecel := cfgStopDecel; END_IF
END_SET
END_PROPERTY

PROPERTY PUBLIC cfgHaltDecel : LREAL
GET
cfgHaltDecel := _haltDecel;
END_GET
SET
IF cfgHaltDecel > 0.0 THEN _haltDecel := cfgHaltDecel; END_IF
END_SET
END_PROPERTY

PROPERTY PUBLIC cfgVelocityOverride : LREAL
GET
cfgVelocityOverride := _velocityOverride;
END_GET
SET
IF cfgVelocityOverride >= 0.0 AND cfgVelocityOverride <= 100.0 THEN
    _velocityOverride := cfgVelocityOverride;
END_IF
END_SET
END_PROPERTY

PROPERTY PUBLIC cfgAccelOverride : LREAL
GET
cfgAccelOverride := _accelOverride;
END_GET
SET
IF cfgAccelOverride >= 0.0 AND cfgAccelOverride <= 100.0 THEN
    _accelOverride := cfgAccelOverride;
END_IF
END_SET
END_PROPERTY

PROPERTY cfgDeviceName : STRING
GET
cfgDeviceName := _deviceName;
END_GET
SET
_deviceName := cfgDeviceName;
END_SET
END_PROPERTY

// Linear vs rotary - for HMI unit display only (NC has no kinematic type).
PROPERTY PUBLIC cfgAxisType : E_Axis_UnitType
GET
cfgAxisType := _axisType;
END_GET
SET
_axisType := cfgAxisType;
END_SET
END_PROPERTY

// Engineering unit label for position (e.g. 'mm', 'deg', 'rev'). HMI shows
// velocity as this + '/s'.
PROPERTY PUBLIC cfgUnit : STRING
GET
cfgUnit := _unit;
END_GET
SET
_unit := cfgUnit;
END_SET
END_PROPERTY

// TRUE = the NC axis is configured as a modulo axis. Metadata only (the NC carries no
// modulo flag in the cyclic image); drives whether the HMI shows the modulo position
// (ModuloActPos) or the accumulated ActPos. Orthogonal to cfgAxisType.
PROPERTY PUBLIC cfgIsModulo : BOOL
GET
cfgIsModulo := _isModulo;
END_GET
SET
_isModulo := cfgIsModulo;
END_SET
END_PROPERTY

END_FUNCTION_BLOCK

// ---- POUs/FBs/fb_HmiEventLog.TcPOU
FUNCTION_BLOCK fb_HmiEventLog
(* fb_HmiEventLog

   Buffered HMI event log — a fixed-size RING of recent log lines plus a monotonic sequence number,
   made to be republished in an MQTT transaction group (or any snapshot transport). The HMI backend
   DRAINS the ring by sequence number, so every event is captured regardless of the publish rate —
   unlike sampling a single "current status" string, which silently drops any change shorter than one
   publish period.

   Each slot holds "<seq>|<sev>|<message>" (sev: I=info, W=warning, E=error); slot index = seq MOD
   cRING_SIZE. Usage:
     _log.Info('Auto sequence started');   // or .Warn(...) / .Fault(...) / .Push('I', msg)
   then register stsSequence + stsRingBuffer[0..N-1] into the HMI publish group. The backend keeps a
   "last drained seq" and appends every slot whose seq is newer, so nothing is lost between snapshots
   as long as the ring is larger than the burst between two snapshots (16 covers a 1 s group period).
*)

VAR CONSTANT
	cRING_SIZE		: DINT := 16;	// ring slots; keep the stsRingBuffer array bound below in sync
END_VAR

VAR
	_sequence		: DINT;
END_VAR

VAR_OUTPUT
	stsSequence		: DINT;								// monotonic high-water sequence (also total logged)
	stsRingBuffer	: ARRAY[0..15] OF STRING(120);		// last cRING_SIZE entries, each "<seq>|<sev>|<message>"
	stsRingSize		: DINT := 16;						// exposed so the reader need not hard-code the size
END_VAR

// No cyclic logic — the ring is driven entirely by the Push / Info / Warn / Fault methods.

METHOD PUBLIC Fault : BOOL
VAR_INPUT
	inpMessage		: STRING;
END_VAR
Push('E', inpMessage);
END_METHOD

METHOD PUBLIC Info : BOOL
VAR_INPUT
	inpMessage		: STRING;
END_VAR
Push('I', inpMessage);
END_METHOD

// Append one entry to the ring: "<seq>|<sev>|<message>" at slot (seq MOD cRING_SIZE).
METHOD PUBLIC Push : BOOL
VAR_INPUT
	inpSeverity		: STRING;	// 'I' | 'W' | 'E'
	inpMessage		: STRING;
END_VAR
VAR
	entry			: STRING(120);
END_VAR
_sequence := _sequence + 1;
entry := DINT_TO_STRING(_sequence);
entry := CONCAT(entry, '|');
entry := CONCAT(entry, inpSeverity);
entry := CONCAT(entry, '|');
entry := CONCAT(entry, inpMessage);
stsRingBuffer[_sequence MOD cRING_SIZE] := entry;
stsSequence := _sequence;
END_METHOD

METHOD PUBLIC Warn : BOOL
VAR_INPUT
	inpMessage		: STRING;
END_VAR
Push('W', inpMessage);
END_METHOD

END_FUNCTION_BLOCK

// ---- POUs/FBs/fb_Machine.TcPOU
FUNCTION_BLOCK fb_Machine

VAR_INPUT
	inpReset				: BOOL;		// IO Reset button
	inpStop					: BOOL;		// IO Stop button
	inpStart				: BOOL;		// IO Start button
	inpStartedFeedback		: BOOL;		// State feedback from state machine
	inpBypassInterlocks		: BOOL;		// IO interlock bypass switch
	inpAuto					: BOOL;		// IO Auto 
	inpPause				: BOOL;		// IO Pause button
	inpPausedFeedback		: BOOL;		// State feedback from state machine
	inpSafetyPowerOn		: BOOL;		// Feedback from safety controller
	inpSafetyFaultActive	: BOOL;		// Feedback from safety controller
	inpSafetyFaultDelay		: BOOL;		// Feedback from safety controller
	inpSafetyResetButton	: BOOL;		// IO safety reset
END_VAR

VAR
	HMI					: ST_Machine_HMI_Interface;
	_faultMonitor		: fb_FaultMonitor;
	eventLogger 		: FB_tcEventLogger;
	firstScanTOF	  	: TOF;
	_clearLogs			: BOOL;
	_cmdStop			: BOOL;
	_cmdStart			: BOOL;
	_reset				: BOOL;
	_stop				: BOOL;
	_start				: BOOL;
	_auto				: BOOL;
	_pause				: BOOL;
	_interlockbypass	: BOOL;
	_safetyPowerOn		: BOOL;
	_safetyFaultActive	: BOOL;
	_safetyFaultDelay	: BOOL;
	transSafetyReset	: R_TRIG;
	hostname		  	: fb_gethostname;
	_firstScan			: BOOL := TRUE;
	// --- machine identity = the IPC hostname (2026-09-20) ---
	_machineName		: T_MaxString;	// set once FB_GetHostName has answered; empty before that
	_hostnameRetry		: TON;			// re-arms the lookup while it keeps failing (cold restart: system service not ready yet)
	_hostnameAttempts	: UDINT;		// diagnostic: how many asks it took
	_identityLogged		: BOOL;
	_clearLogTrig		: BOOL;
	MachineState		: fb_Dev_Machine(cfgDeviceName := 'Machine', cfgEnable := TRUE, cfgInitEventClass :=TRUE,);
	myUPS 				: FB_S_UPS_BAPI;
	writePersistent	  	: fb_WritePersistentData;
	writePersTrig	  	: BOOL;
	_hasUPS				: BOOL;
	_hbTimer			: TON;		// 500ms heartbeat generator (HMI frozen-data watchdog)
	_heartbeat			: BOOL;		// toggled square wave published to HMI.stsHeartBeat
END_VAR

VAR_OUTPUT
	stsAuto					: BOOL;
	stsInterlocksBypassed	: BOOL;
	stsFirstScan			: BOOL;
	stsMachineName			: T_MaxString;
	stsIdentityValid		: BOOL;		// TRUE once stsMachineName holds the IPC hostname
	stsStarted				: BOOL;
	stsFaultActive			: BOOL;
	outStop					: BOOL;
	outReset				: BOOL;
	outStart				: BOOL;
END_VAR

firstScanTOF(IN:=_clearLogTrig,PT:=T#20ms);

//Machine identity = the IPC hostname, nothing else. FB_GetHostName is one ADS
//call to the local system service; right after a cold restart it can fail or
//time out, and the old one-shot on the first scan then left the name empty for
//good, and everything keyed on the machine name never started. Ask until it answers.
hostname(sNetID:='', tTimeout:=T#2S);
IF hostname.bExecute AND NOT hostname.bBusy THEN
	// request finished: the result or the error is in
	hostname.bExecute := FALSE;
	IF NOT hostname.bError AND hostname.sHostName <> '' THEN
		_machineName := hostname.sHostName;
	END_IF
END_IF
_hostnameRetry(IN := (_machineName = '') AND NOT hostname.bExecute AND NOT hostname.bBusy, PT := T#1S);
IF (_firstScan OR _hostnameRetry.Q) AND _machineName = '' AND NOT hostname.bExecute THEN
	hostname.bExecute := TRUE;
	_hostnameAttempts := _hostnameAttempts + 1;
END_IF
IF _machineName <> '' AND NOT _identityLogged THEN
	_identityLogged := TRUE;
	ADSLOGSTR(ADSLOG_MSGTYPE_HINT OR ADSLOG_MSGTYPE_LOG,
		CONCAT(CONCAT('Machine identity acquired after ', UDINT_TO_STRING(_hostnameAttempts)), ' attempt(s): %s'), _machineName);
END_IF

// Run UPS
IF _hasUPS THEN
	myUPS(sNetID :='',
			iPLCPort:=851,
		  tTimeout := DEFAULT_ADS_TIMEOUT,
		  eUPSMode := eSUPS_WrPersistData_Shutdown,
		  ePersistentMode := SPDM_2PASS,tRecoverTime := T#3S);
	writePersistent(NETID:='', PORT := 851, START:= writePersTrig,TMOUT := DEFAULT_ADS_TIMEOUT);
END_IF

//Run global fault monitor	  
_faultMonitor();

// Interlock Bypass

_interlockBypass := inpBypassInterlocks;

//Send out Reset oneshot if reset is triggered from HMI, safety button, or method
transSafetyReset(CLK:=inpSafetyResetButton);
IF transSafetyReset.q OR HMI.inpReset OR _reset OR inpReset THEN
	HMI.inpReset 	:= FALSE;
	_reset			:= FALSE;
	outReset	 	:= TRUE;
	IF _stop THEN
		_stop := FALSE;
	END_IF
ELSE
	outReset 		:= FALSE;
END_IF

IF HMI.inpManual THEN
	HMI.inpManual 	:= FALSE;
	_auto 			:= FALSE;
END_IF

IF HMI.inpAuto OR inpAuto THEN
	HMI.inpAuto 	:= FALSE;
	_auto			:= TRUE;
END_IF

IF HMI.inpStart OR _cmdStart THEN
	HMI.inpStart := FALSE;
	_cmdStart	 := FALSE;
	outStart	 := TRUE;
ELSE
	outStart	:= FALSE;
END_IF

IF HMI.inpStop OR inpStop OR _cmdStop THEN
	HMI.inpStop	:= FALSE;
	_cmdStop	:= FALSE;
	_start		:= FALSE;
	_stop		:= TRUE;
END_IF

IF HMI.inpClearMachineLog OR _clearLogs THEN
	HMI.inpClearMachineLog := FALSE;
	_clearLogs		:= FALSE;
	_clearLogTrig	:= TRUE;
END_IF

IF firstScanTOF.Q THEN
	_clearLogTrig	:= FALSE;
	eventLogger.ClearLoggedEvents(0);
END_IF

HMI.stsMachineName			:= _machineName;
HMI.stsInAuto				:= _auto;
HMI.stsInManual				:= NOT(_auto);
HMI.stsInterlockBypassed	:= _interlockbypass;
HMI.stsPaused				:= inpPausedFeedback;
HMI.stsStarted				:= inpStartedFeedback;
HMI.stsStopped				:= _stop;

// HMI heartbeat: 500ms on / 500ms off square wave the web HMI watches to detect frozen data
// end-to-end (PLC stopped / stale reads) even while the transport still reads OK.
_hbTimer(IN := NOT _hbTimer.Q, PT := T#500MS);
IF _hbTimer.Q THEN
	_heartbeat := NOT _heartbeat;
END_IF
HMI.stsHeartBeat			:= _heartbeat;

_safetyPowerOn				:= inpSafetyPowerOn;
_safetyFaultActive			:= inpSafetyFaultActive;
_safetyFaultDelay			:= inpSafetyFaultDelay;

MachineState(inpAuto := _auto, inpReset := outReset, inpInterlockbypass := _interlockbypass, start:=_start, stop:=_stop
			, SafetyPowerOn:= _safetyPowerOn, SafetyFaultActive:=_safetyFaultActive, faultMonitor :=ADR(_faultMonitor));

stsAuto						:= _auto;
stsInterlocksBypassed		:= _interlockbypass;
stsFirstScan				:= _firstScan;
stsMachineName				:= _machineName;
stsIdentityValid			:= _machineName <> '';
stsStarted					:= inpStartedFeedback;
outStop						:= _stop;
stsFaultActive				:= _faultMonitor.stsFaultActive;

PROPERTY cfgHasUPS : bool
GET
cfgHasUPS := _hasUPS;
END_GET
SET
_hasUPS := cfgHasUPS;
END_SET
END_PROPERTY

METHOD cmdClearLogs : BOOL
VAR_INPUT
END_VAR
_clearLogs := TRUE;
END_METHOD

METHOD cmdExportEventLogs : BOOL
VAR_INPUT
	filePath : T_MaxString;
END_VAR
VAR
	exportSettings : FB_TcEventCsvExportSettings;
END_VAR
exportSettings.sDelimiter := ',';
eventLogger.ExportLoggedEvents(sFilename := filePath, ipExportSettings:=exportSettings);
END_METHOD

METHOD cmdReset : BOOL
VAR_INPUT
END_VAR
_reset := TRUE;
END_METHOD

METHOD cmdStart : BOOL
VAR_INPUT
END_VAR
_cmdStart := TRUE;
END_METHOD

METHOD cmdStop : BOOL
VAR_INPUT
END_VAR
_cmdStop := TRUE;
END_METHOD

PROPERTY faultMonitor : POINTER TO fb_faultmonitor
GET
faultMonitor := ADR(_faultMonitor);
END_GET
END_PROPERTY

//FB_Init is always available implicitly and it is used primarily for initialization.
//The return value is not evaluated. For a specific influence, you can also declare the
//methods explicitly and provide additional code there with the standard initialization
//code. You can evaluate the return value.
METHOD FB_Init: BOOL
VAR_INPUT
    bInitRetains: BOOL; // TRUE: the retain variables are initialized (reset warm / reset cold)
    bInCopyCode: BOOL;  // TRUE: the instance will be copied to the copy code afterward (online change)   
	hasUPS		: BOOL;
END_VAR
THIS^._hasUPS := hasUPS;
END_METHOD

METHOD firstScanComplete : BOOL
VAR_INPUT
END_VAR
_firstScan := FALSE;
END_METHOD

END_FUNCTION_BLOCK

// ---- POUs/FBs/fb_PID_Clamping.TcPOU
FUNCTION_BLOCK fb_PID_Clamping
VAR_INPUT
    inpSP               : LREAL;
    inpPV               : LREAL;
    inpManualValue      : LREAL;
    inpEnable           : BOOL;
    inpPIDReset         : BOOL;
    cfgKp               : LREAL;
    cfgTn               : LREAL;
    cfgTv               : LREAL;
    cfgOutMin           : LREAL := 0.0;
    cfgOutMax           : LREAL := 350.0;
    cfgCycleTime        : LREAL := 0.01;
    cfgOutputFilterAlpha: LREAL := 0.4;
    cfgDerivFilterN     : LREAL := 8.0;
    cfgPvRateWindow     : LREAL := 20.0;
    cfgCoolingMode      : BOOL := FALSE;
END_VAR
VAR_OUTPUT
    stsOut              : LREAL;
    stsAuto             : BOOL;
END_VAR
VAR
    _integral           : LREAL;
    _p                  : LREAL;
    _i                  : LREAL;
    _d                  : LREAL;
    _pvRate             : LREAL;
    _pvWindowAgo        : LREAL;
    _windowTimer        : LREAL;
    _error              : LREAL;
    _outRaw             : LREAL;
    _outClamped         : LREAL;
    _wasAuto            : BOOL;
END_VAR

// Reset clears accumulated controller state only. It must NOT force the output
// to 0, otherwise it would override the manual pass-through below when reset is
// held while the block is disabled.
IF inpPIDReset THEN
    _integral    := 0.0;
    _pvWindowAgo := inpPV;
    _windowTimer := 0.0;
    _d           := 0.0;
    _wasAuto     := FALSE;
END_IF

// Error sign depends on mode. Heating: drive output up when PV is below SP.
// Cooling: drive output up when PV is above SP (reverse acting).
IF cfgCoolingMode THEN
    _error := inpPV - inpSP;
ELSE
    _error := inpSP - inpPV;
END_IF

// Disabled: pass the manual value straight through (transparent insert) and
// preload the integral so the first auto scan resumes from the manual value.
IF NOT inpEnable THEN
    _outClamped := LIMIT(cfgOutMin, inpManualValue, cfgOutMax);
    stsOut      := _outClamped;
    stsAuto     := FALSE;
    _wasAuto     := FALSE;
    _pvWindowAgo := inpPV;
    _windowTimer := 0.0;
    _d           := 0.0;
    _p           := cfgKp * _error;
    _integral    := _outClamped - _p;
    RETURN;
END_IF

stsAuto := TRUE;

// On transfer into auto, seed the rate window and clear the filtered derivative
// so the first scan sees no PV step and no carried-over derivative state.
IF NOT _wasAuto THEN
    _pvWindowAgo := inpPV;
    _windowTimer := 0.0;
    _d           := 0.0;
    _wasAuto     := TRUE;
END_IF

_p := cfgKp * _error;

IF cfgTn > 0.0 THEN
    IF (_outClamped >= cfgOutMax AND _error > 0.0) OR
       (_outClamped <= cfgOutMin AND _error < 0.0) THEN
        ;
    ELSE
        _integral := _integral + (cfgKp / cfgTn) * _error * cfgCycleTime;
    END_IF
    _i := _integral;
ELSE
    _i := 0.0;
END_IF

// Derivative on measurement (PV), first-order filtered.
//
// Acting on the change in PV (not error) avoids a derivative kick when the
// setpoint moves and keeps the sign convention explicit. The filter is the
// backward-Euler discretization of  Kp*Tv*s / (1 + (Tv/N)*s), with divisor N:
// large N -> near-raw difference, small N -> heavier smoothing. It rejects the
// per-tick spikes produced by the 0.1 degC PV quantization so the term tracks
// the genuine temperature trend instead of chattering on each digit step.
//
// Sign: a rising PV must raise output in cooling mode (anticipatory fan
// spin-up) and lower it in heating mode.
IF cfgTv > 0.0 AND cfgDerivFilterN > 0.0 THEN
    // PV is quantized to 0.1 degC and changes slowly (~0.1 degC / 30 s), so a
    // scan-to-scan difference is 0.0 on almost every scan. Measure the change
    // over a fixed window instead and divide by the elapsed window time to get
    // a true degC/s rate. _pvRate updates once per window and holds between
    // updates; the process is far slower than the window and the derivative
    // filter below smooths the steps.
    _windowTimer := _windowTimer + cfgCycleTime;
    IF _windowTimer >= cfgPvRateWindow THEN
        IF cfgCoolingMode THEN
            _pvRate := (inpPV - _pvWindowAgo) / _windowTimer;
        ELSE
            _pvRate := (_pvWindowAgo - inpPV) / _windowTimer;
        END_IF
        _pvWindowAgo := inpPV;
        _windowTimer := 0.0;
    END_IF
    _d := (cfgTv / (cfgTv + cfgDerivFilterN * cfgCycleTime)) * _d
        + (cfgKp * cfgTv * cfgDerivFilterN / (cfgTv + cfgDerivFilterN * cfgCycleTime)) * _pvRate;
ELSE
    _d := 0.0;
END_IF

_outRaw     := _p + _i + _d;
_outClamped := LIMIT(cfgOutMin, _outRaw, cfgOutMax);

// Smooth the output
stsOut := stsOut + cfgOutputFilterAlpha * (_outClamped - stsOut);

END_FUNCTION_BLOCK

// ---- POUs/FBs/fb_RampGenerator.TcPOU
FUNCTION_BLOCK fb_RampGenerator
VAR_INPUT
    inpSPRequest    : LREAL;    (* Requested Setpoint value *)
    inpRampTime     : TIME;     (* Total desired time for the ramp (e.g., T#5s, T#250ms).
                                   If T#0s or less, output jumps immediately. *)
    cfgScanRate     : TIME;     (* Scan rate (cycle time) of the task calling this FB instance
                                   (e.g., T#1ms, T#10ms). Must be greater than T#0s. *)
END_VAR
VAR_OUTPUT
    stsRamp         : LREAL;    (* Current ramped output value *)
	stsRampActive	: BOOL;
END_VAR
VAR
    // Internal state variables
    _lastSPRequest  : LREAL;    (* Stores the previous SP request to detect changes *)
    _startValue     : LREAL;    (* Value of stsRamp when the ramp started *)
    _targetValue    : LREAL;    (* Target value (inpSPRequest) for the current ramp *)
    _increment      : LREAL;    (* Amount to add/subtract from stsRamp each scan cycle *)
    _scanCounter    : UDINT;    (* Counts scans elapsed during the current ramp *)
    _totalScans     : UDINT;    (* Total number of scans required for the complete ramp *)
    _isRamping      : BOOL := FALSE; (* TRUE if a ramp is currently in progress *)
    _firstScan      : BOOL := TRUE;  (* Flag for first scan initialization *)

    // Internal calculation variables
    _rampTimeSeconds : LREAL;   (* Calculated ramp time in seconds *)
    _scanRateSeconds : LREAL;   (* Calculated scan rate in seconds *)
END_VAR
VAR CONSTANT
    MILLISECONDS_TO_SECONDS : LREAL := 1000.0; (* Conversion factor *)
    ZERO_LREAL              : LREAL := 0.0;    (* Constant for zero LREAL *)
END_VAR

// --- Initialization on the first scan cycle ---
// On the very first call after instantiation or reset, initialize internal states.
IF _firstScan THEN
    stsRamp         := inpSPRequest;        // Initialize output to the initial request
    _lastSPRequest  := inpSPRequest;        // Initialize last request tracking
    _targetValue    := inpSPRequest;        // Initialize target value
    _startValue     := inpSPRequest;        // Initialize start value
    _isRamping      := FALSE;               // Not ramping initially
    _scanCounter    := 0;
    _totalScans     := 0;
    _increment      := ZERO_LREAL;
    _firstScan      := FALSE;               // Clear the first scan flag for subsequent calls
END_IF

// --- Check for Setpoint Change ---
// Detect if the external request has changed since the last scan cycle.
IF inpSPRequest <> _lastSPRequest THEN
    // A new ramp needs to be started or the target needs immediate update.
    _targetValue    := inpSPRequest;   // Store the new target value
    _startValue     := stsRamp;        // The ramp starts from the current output value

    // --- Calculate Ramp Parameters ---
    // Convert TIME inputs to LREAL seconds for calculation.
    // Uses the native TIME_TO_LREAL function (converts TIME to LREAL milliseconds)
    // and divides by 1000.0 to get seconds. Requires Standard.lib (usually included).
    _rampTimeSeconds := TIME_TO_LREAL(inpRampTime) / MILLISECONDS_TO_SECONDS;
    _scanRateSeconds := TIME_TO_LREAL(cfgScanRate) / MILLISECONDS_TO_SECONDS;

    // Check for valid positive ramp time and scan rate. Scan rate must be positive.
    IF _rampTimeSeconds > ZERO_LREAL AND _scanRateSeconds > ZERO_LREAL THEN
        // Calculate the total number of scan cycles required for the ramp duration.
        // LREAL_TO_UDINT truncates; for very precise timing, consider rounding logic if needed.
        _totalScans := LREAL_TO_UDINT(_rampTimeSeconds / _scanRateSeconds);

        IF _totalScans > 0 AND _targetValue <> _startValue THEN
            // Calculate the change in value required per scan cycle.
            _increment := (_targetValue - _startValue) / UDINT_TO_LREAL(_totalScans);
            _scanCounter := 0;      // Reset the scan counter for the new ramp
            _isRamping := TRUE;     // Set the flag indicating ramp is active
        ELSE
            // Ramp time is shorter than one scan cycle, total scans is zero,
            // or start value already equals target value. Jump directly.
            stsRamp := _targetValue;
            _isRamping := FALSE;
            _scanCounter := 0;
            _totalScans := 0;
            _increment := ZERO_LREAL;
        END_IF
    ELSE
        // Ramp time is zero/negative or scan rate is invalid (zero/negative). Jump directly.
        stsRamp := _targetValue;
        _isRamping := FALSE;
        _scanCounter := 0;
        _totalScans := 0;
        _increment := ZERO_LREAL;
    END_IF

    // Update the last tracked SP request AFTER calculations are done based on the change.
    _lastSPRequest := inpSPRequest;

// --- Continue Active Ramp ---
ELSIF _isRamping THEN
    // If the Setpoint Request hasn't changed, continue the current ramp if one is active.
    IF _scanCounter < _totalScans THEN
        // Increment/decrement the ramp value by the calculated step.
        stsRamp := stsRamp + _increment;
        _scanCounter := _scanCounter + 1;

        // Check if the ramp is now complete (reached or passed target) on this scan.
        // This check prevents overshoot/undershoot due to floating point inaccuracies
        // and ensures the ramp stops exactly at the target value.
        IF _scanCounter >= _totalScans OR
           (_increment > ZERO_LREAL AND stsRamp >= _targetValue) OR
           (_increment < ZERO_LREAL AND stsRamp <= _targetValue) THEN

            stsRamp := _targetValue; // Set final value exactly
            _isRamping := FALSE;     // Mark ramp as finished
            // Optional: _scanCounter := _totalScans; // Ensure counter reflects completion state
        END_IF
    ELSE
        // Safeguard: If ramp flag is somehow still true but counter is already >= total, fix state.
        stsRamp := _targetValue;
        _isRamping := FALSE;
    END_IF
END_IF

stsRampActive := _isRamping;

END_FUNCTION_BLOCK

// ---- POUs/FBs/fb_SampleBuffer.TcPOU
(* fb_SampleBuffer

   Sensor-agnostic oversampling ring buffer. Captures the N-sample oversample
   block delivered by a Beckhoff oversampling terminal each PLC scan (1 ms
   scan) into a long ring buffer that an external ADS reader (the chart
   engine) can poll at its own slower cadence without losing samples.

   Works for any terminal that produces a block of 32-bit samples per scan:
     - ELM3602-0002 accelerometer (raw INT32 ADC counts, 50 kHz / 50x)
     - EL5101-0011 encoder (oversampled position counter, for order tracking)
   The FB doesn't interpret the samples — it just rings them. Scaling /
   unwrapping / FFT happen downstream in the engine, so a DINT ring is used
   regardless of what the counts mean (encoder UDINT counters are bit-
   compatible; map them as DINT in the process image and unwrap in Python).

   The engine's actual fast-loop period on a reference test-stand config measures
   ~80 ms (89-signal batch + 2x 16 KB ring reads + asyncio.sleep(33 ms)), so
   the ring consumes ~4000 samples per tick. cRING_SIZE = 8192 gives ~164 ms
   of buffer — absorbing both the slow first tick (extra slow + test-panel
   reads, ~115 ms) and transient ADS jitter without overwriting unread samples.

   Reader contract:
     - stsTotalSamples is monotonic across PLC restarts of this FB (never wraps
       for ~12,000 years at 50 kHz). The reader stores its last-seen value;
       delta := stsTotalSamples - lastSeen tells the reader how many new samples
       arrived since the previous read.
     - If delta > stsRingSize the reader has fallen behind further than the
       ring can hold — older samples have been overwritten. Detection and
       handling (gap-marker, drop window, log) live on the reader side.
     - To extract the last N := MIN(delta, stsRingSize) samples in chrono
       order, read backward from ((stsWriteIdx - 1) MOD stsRingSize) for N
       slots, then reverse — or read the whole stsRingBuffer once and slice.

   For synchronous multi-channel work (e.g. order tracking pairs an accel
   instance with an encoder instance): instantiate one FB per signal in the
   same task. All instances advance stsTotalSamples in lockstep (+cBLOCK_SIZE
   per scan), so the reader aligns channels by total-sample index.
*)
FUNCTION_BLOCK fb_SampleBuffer

VAR CONSTANT
	cRING_SIZE		: UDINT := 8192;	// ~164 ms of buffer at 50 kHz; absorbs slow first tick + ADS jitter
	cBLOCK_SIZE		: UDINT := 50;		// oversample factor at 1 ms scan (ELM3602 / EL5101 50x)
END_VAR

VAR_INPUT
	inpRawBlock		: ARRAY [0..49] OF DINT;	// one oversample frame (accel block or encoder block)
	inpEnable		: BOOL := TRUE;
END_VAR

VAR_OUTPUT
	stsRingBuffer	: ARRAY [0..8191] OF DINT;	// raw samples; reader uses stsTotalSamples to compute the newest-sample slot
	stsTotalSamples	: ULINT;					// monotonic count of samples ever written; never wraps in practice
	stsWriteIdx		: UDINT;					// next slot to write into; ((stsWriteIdx - 1) MOD cRING_SIZE) is newest
	stsRingSize		: UDINT := 8192;			// exposed for the reader so it doesn't have to hard-code
	stsBlockSize	: UDINT := 50;
END_VAR

VAR
	_writeIdx		: UDINT;
END_VAR

IF NOT inpEnable THEN
	RETURN;
END_IF

BufferSamples();

stsWriteIdx := _writeIdx;

(* Append the oversample frame into the ring and advance the monotonic
   sample counter. Wrapping is per-sample (not per-block) so reader logic
   doesn't need to special-case partial-block wraps. *)
METHOD BufferSamples : BOOL
VAR
	i : UDINT;
END_VAR
FOR i := 0 TO cBLOCK_SIZE - 1 DO
	stsRingBuffer[_writeIdx] := inpRawBlock[i];
	_writeIdx := (_writeIdx + 1) MOD cRING_SIZE;
END_FOR

stsTotalSamples := stsTotalSamples + cBLOCK_SIZE;
END_METHOD

END_FUNCTION_BLOCK

// ---- POUs/FBs/fb_TimeAverage.TcPOU
FUNCTION_BLOCK fb_TimeAverage
VAR_INPUT
    inpSignal         : LREAL;         // The input signal to be averaged
    inpSampleTime     : TIME := T#10MS; // The cycle time of the task calling this FB (e.g., 10ms)
    inpAverageTime    : TIME := T#1s;   // The desired time window for the average (e.g., 1s)
END_VAR
VAR_OUTPUT
    outAverage        : LREAL;         // The calculated average value over the specified time
END_VAR
VAR
    rSum            : LREAL;        // Use LREAL for the sum to avoid precision loss with many additions
    nSampleCount    : DINT;         // Counter for the number of samples collected
    nMaxSamples     : DINT;         // The total number of samples required for the averaging period
    bInitialize     : BOOL := TRUE; // Flag to initialize on the first scan
END_VAR

IF bInitialize THEN
    // Ensure tSampleTime is not zero to prevent division by zero error.
    IF inpSampleTime > T#0S THEN
        // Calculate the number of samples needed to fill the averaging time window.
        // We convert TIME to DINT (in nanoseconds) for the calculation.
        nMaxSamples := TIME_TO_DINT(inpAverageTime) / TIME_TO_DINT(inpSampleTime);
    ELSE
        // If sample time is zero, set max samples to 1 to avoid errors.
        nMaxSamples := 1;
    END_IF;
    
    // Reset internal variables to start a fresh calculation
    rSum := 0.0;
    nSampleCount := 0;
    
    // Initialization is complete.
    bInitialize := FALSE;
END_IF

// Accumulate the signal value and increment the sample counter in every scan.
nSampleCount := nSampleCount + 1;
rSum := rSum + inpSignal;

// Check if the required number of samples for the averaging period has been collected.
IF nSampleCount >= nMaxSamples THEN
    // Calculate the average value.
    // Check nSampleCount to be safe, although it should equal nMaxSamples here.
    IF nSampleCount > 0 THEN
        outAverage := rSum / nSampleCount;
    END_IF;
    
    // Reset the sum and counter to begin the next averaging window.
    rSum := 0.0;
    nSampleCount := 0;
END_IF;

END_FUNCTION_BLOCK

// ---- POUs/FC/F_AddToArray_String.TcPOU
FUNCTION F_AddToArray_String : BOOL
VAR_INPUT
    value : STRING;            // String to add
    maxSize : DINT;           // Maximum array capacity
END_VAR
VAR_IN_OUT
    arr : ARRAY[*] OF STRING; // Array of strings
END_VAR
VAR
    currentSize : DINT := 0;
    i : DINT;
END_VAR

F_AddToArray_String := FALSE;

// Find current size by looking for first empty string
FOR i := 1 TO UPPER_BOUND(arr, 1) DO
    IF arr[i] = '' THEN
        currentSize := i;
        EXIT;
    END_IF
    // If we reach the end without finding empty string
    IF i = UPPER_BOUND(arr, 1) THEN
        currentSize := i + 1;
    END_IF
END_FOR

// Check if there's space to add
IF currentSize >= maxSize OR currentSize > UPPER_BOUND(arr, 1) THEN
    RETURN;
END_IF

// Add the string
arr[currentSize] := value;
F_AddToArray_String := TRUE;

END_FUNCTION

// ---- POUs/FC/F_RemoveFromArray_String.TcPOU
FUNCTION F_RemoveFromArray_String : DINT
VAR_INPUT
    value : STRING;            // String to remove
    maxSize : DINT;           // Maximum array capacity
END_VAR
VAR_IN_OUT
    arr : ARRAY[*] OF STRING; // Array of strings
END_VAR
VAR
    currentSize : DINT := 0;
    i : DINT;
    foundPos : DINT := -1;    // -1 indicates not found
END_VAR

// Find current size and position of value
FOR i := 1 TO UPPER_BOUND(arr, 1) DO
    IF arr[i] = '' THEN
        currentSize := i;
        EXIT;
    END_IF
    IF arr[i] = value AND foundPos = -1 THEN
        foundPos := i;
    END_IF
    // If we reach the end without finding empty string
    IF i = UPPER_BOUND(arr, 1) THEN
        currentSize := i + 1;
    END_IF
END_FOR

// If value wasn't found or array is empty, return
IF foundPos = -1 OR currentSize = 0 THEN
    RETURN;
END_IF

// Shift elements up to fill the gap
FOR i := foundPos TO currentSize - 2 DO
    arr[i] := arr[i + 1];
END_FOR

// Clear the last element
arr[currentSize - 1] := '';

// Return the position where the value was found
F_RemoveFromArray_String := foundPos;

END_FUNCTION
